Fanuc KAREL source: KT00550.KL

PROGRAM KT00550
%NOLOCKGROUP
VAR
  P1: JOINTPOS
  P2: JOINTPOS
  OUT: XYZWPR
BEGIN
  OUT = P1 : P2
END KT00550
